(* IEC 61131-3 sources: PLC-Static-Analysis/modules/plc-rules/src/test/resources/PLCA-L012, 2 files *)

(* ---- compliant.st ---- *)
PROGRAM P_L012ok
VAR
    nInt : INT;
    nInt2 : INT;
    nByte : BYTE;
    nDint : DINT;
    nRange : INT(0..10);
    sName : STRING(4);
    q : BOOL;
END_VAR
q := nInt < 0;
q := nByte >= 255;
q := nInt + nInt2 > 32767;
q := nRange > 9;
q := sName = 'ABCD';
q := nDint > 2147483646;
END_PROGRAM

(* ---- noncompliant.st ---- *)
PROGRAM P_L012
VAR
    nUsint : USINT;
    nByte : BYTE;
    nUint : UINT;
    nSint : SINT;
    nRange : INT(0..10);
    sName : STRING(4);
    b : BOOL;
    q : BOOL;
END_VAR
IF nUsint < 0 THEN // PLCA-L012
    q := TRUE;
END_IF
q := nByte > 255; // PLCA-L012
q := nUint >= 0; // PLCA-L012
q := nRange > 10; // PLCA-L012
q := sName = 'TOO_LONG'; // PLCA-L012
q := sName <> 'ALSO_TOO_LONG'; // PLCA-L012
q := nSint = 200 OR b; // PLCA-L012
END_PROGRAM
